// TIA Portal V17 export
// export: Created 2026-11-08T05:50:28.3151889Z, ExportSetting WithDefaults, DisplayName Totally Integrated Automation Portal, DisplayVersion V17, DisplayName TIA Portal Openness, DisplayVersion V17, DisplayName TIA Portal Version Control Interface, DisplayVersion V17, DisplayName STEP 7 Professional, DisplayVersion V17, DisplayName STEP 7 Safety, DisplayVersion V17, DisplayName WinCC Professional, DisplayVersion V17
ORGANIZATION_BLOCK "Main"   // OB1, LAD, ProgramCycle
TITLE = "Main Program Sweep (Cycle)" / Programa principal - Arranque y paro v2
{ S7_Optimized_Access := 'TRUE' }
VERSION : 0.1
// OB1 director: una red por función. Los 3 estilos corren a la vez; el selector de la HMI decide cuál maneja KM1 y los pilotos.
// stored: AutoNumber true, IsIECCheckEnabled false, SetENOAutomatically false
   VAR_INPUT
      Initial_Call : Bool;   // Initial call of this OB
      Remanence : Bool;   // =True, if remanent data are available
   END_VAR
BEGIN

REGION Network 1: MANDO: pulsadores + HMI
   // Une entradas físicas y botones de la HMI.
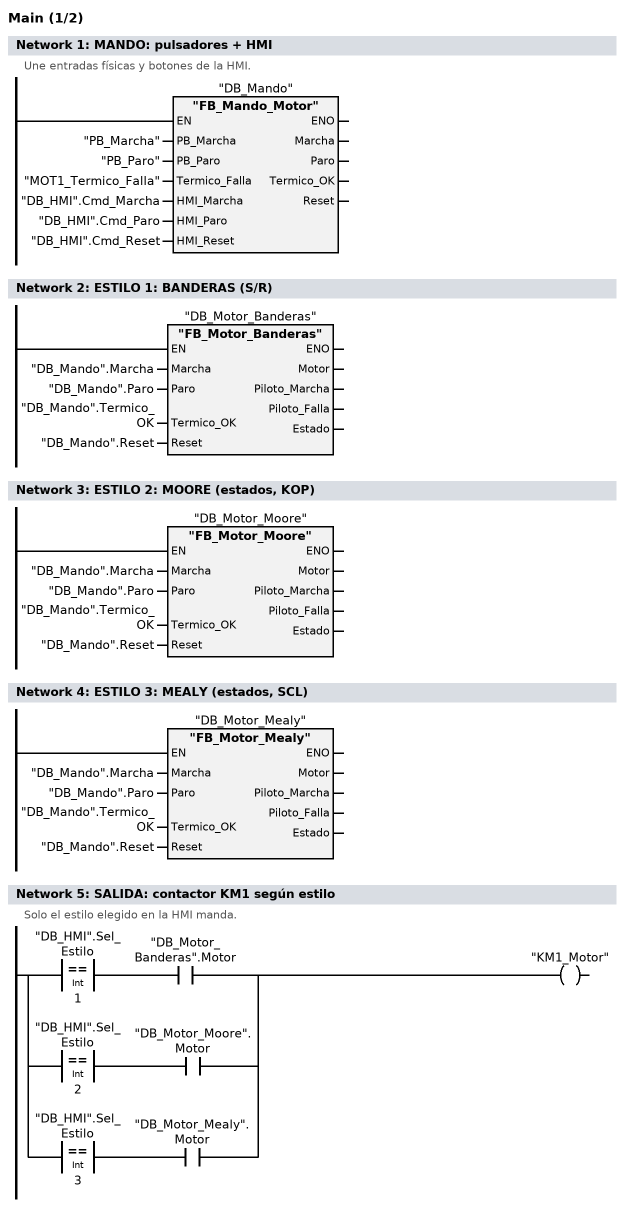
   RUNG wire#powerrail
      "DB_Mando"(PB_Marcha := "PB_Marcha", PB_Paro := "PB_Paro", Termico_Falla := "MOT1_Termico_Falla", HMI_Marcha := "DB_HMI".Cmd_Marcha, HMI_Paro := "DB_HMI".Cmd_Paro, HMI_Reset := "DB_HMI".Cmd_Reset, Marcha =>, Paro =>, Termico_OK =>, Reset =>)
   END_RUNG
   // the same network as SCL:
   "DB_Mando"(PB_Marcha := "PB_Marcha",   // "FB_Mando_Motor"
              PB_Paro := "PB_Paro",
              Termico_Falla := "MOT1_Termico_Falla",
              HMI_Marcha := "DB_HMI".Cmd_Marcha,
              HMI_Paro := "DB_HMI".Cmd_Paro,
              HMI_Reset := "DB_HMI".Cmd_Reset);
END_REGION

REGION Network 2: ESTILO 1: BANDERAS (S/R)
   RUNG wire#powerrail
      "DB_Motor_Banderas"(Marcha := "DB_Mando".Marcha, Paro := "DB_Mando".Paro, Termico_OK := "DB_Mando".Termico_OK, Reset := "DB_Mando".Reset, Motor =>, Piloto_Marcha =>, Piloto_Falla =>, Estado =>)
   END_RUNG
   // the same network as SCL:
   "DB_Motor_Banderas"(Marcha := "DB_Mando".Marcha,   // "FB_Motor_Banderas"
                       Paro := "DB_Mando".Paro,
                       Termico_OK := "DB_Mando".Termico_OK,
                       Reset := "DB_Mando".Reset);
END_REGION

REGION Network 3: ESTILO 2: MOORE (estados, KOP)
   RUNG wire#powerrail
      "DB_Motor_Moore"(Marcha := "DB_Mando".Marcha, Paro := "DB_Mando".Paro, Termico_OK := "DB_Mando".Termico_OK, Reset := "DB_Mando".Reset, Motor =>, Piloto_Marcha =>, Piloto_Falla =>, Estado =>)
   END_RUNG
   // the same network as SCL:
   "DB_Motor_Moore"(Marcha := "DB_Mando".Marcha,   // "FB_Motor_Moore"
                    Paro := "DB_Mando".Paro,
                    Termico_OK := "DB_Mando".Termico_OK,
                    Reset := "DB_Mando".Reset);
END_REGION

REGION Network 4: ESTILO 3: MEALY (estados, SCL)
   RUNG wire#powerrail
      "DB_Motor_Mealy"(Marcha := "DB_Mando".Marcha, Paro := "DB_Mando".Paro, Termico_OK := "DB_Mando".Termico_OK, Reset := "DB_Mando".Reset, Motor =>, Piloto_Marcha =>, Piloto_Falla =>, Estado =>)
   END_RUNG
   // the same network as SCL:
   "DB_Motor_Mealy"(Marcha := "DB_Mando".Marcha,   // "FB_Motor_Mealy"
                    Paro := "DB_Mando".Paro,
                    Termico_OK := "DB_Mando".Termico_OK,
                    Reset := "DB_Mando".Reset);
END_REGION

REGION Network 5: SALIDA: contactor KM1 según estilo
   // Solo el estilo elegido en la HMI manda.
   RUNG wire#powerrail
      { S7_Templates := "SrcType := Int" } EQ_Contact(in1 := "DB_HMI".Sel_Estilo, in2 := 1)
      Contact( "DB_Motor_Banderas".Motor )
      wire#w1
      Coil( "KM1_Motor" )
   END_RUNG
   RUNG wire#powerrail
      { S7_Templates := "SrcType := Int" } EQ_Contact(in1 := "DB_HMI".Sel_Estilo, in2 := 2)
      Contact( "DB_Motor_Moore".Motor )
   END_RUNG wire#w1
   RUNG wire#powerrail
      { S7_Templates := "SrcType := Int" } EQ_Contact(in1 := "DB_HMI".Sel_Estilo, in2 := 3)
      Contact( "DB_Motor_Mealy".Motor )
   END_RUNG wire#w1
   // the same network as SCL:
   "KM1_Motor" := (("DB_HMI".Sel_Estilo = 1) AND "DB_Motor_Banderas".Motor) OR (("DB_HMI".Sel_Estilo = 2) AND "DB_Motor_Moore".Motor) OR (("DB_HMI".Sel_Estilo = 3) AND "DB_Motor_Mealy".Motor);
END_REGION

REGION Network 6: SALIDA: piloto de marcha
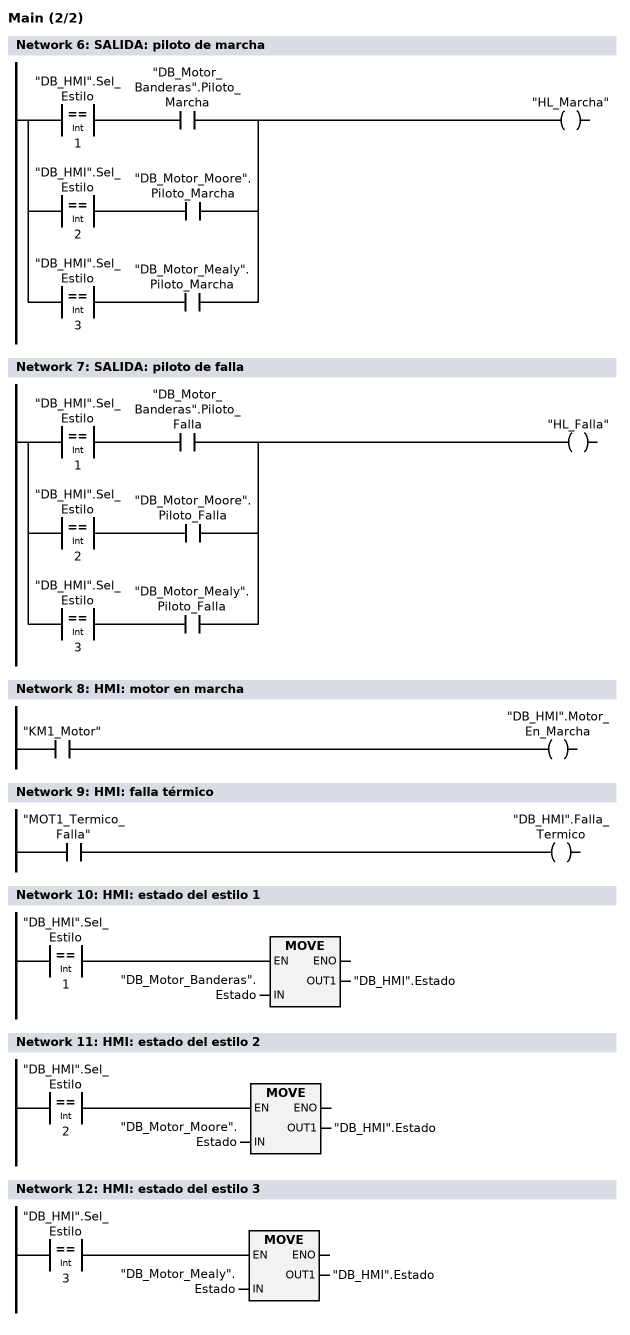
   RUNG wire#powerrail
      { S7_Templates := "SrcType := Int" } EQ_Contact(in1 := "DB_HMI".Sel_Estilo, in2 := 1)
      Contact( "DB_Motor_Banderas".Piloto_Marcha )
      wire#w1
      Coil( "HL_Marcha" )
   END_RUNG
   RUNG wire#powerrail
      { S7_Templates := "SrcType := Int" } EQ_Contact(in1 := "DB_HMI".Sel_Estilo, in2 := 2)
      Contact( "DB_Motor_Moore".Piloto_Marcha )
   END_RUNG wire#w1
   RUNG wire#powerrail
      { S7_Templates := "SrcType := Int" } EQ_Contact(in1 := "DB_HMI".Sel_Estilo, in2 := 3)
      Contact( "DB_Motor_Mealy".Piloto_Marcha )
   END_RUNG wire#w1
   // the same network as SCL:
   "HL_Marcha" := (("DB_HMI".Sel_Estilo = 1) AND "DB_Motor_Banderas".Piloto_Marcha) OR (("DB_HMI".Sel_Estilo = 2) AND "DB_Motor_Moore".Piloto_Marcha) OR (("DB_HMI".Sel_Estilo = 3) AND "DB_Motor_Mealy".Piloto_Marcha);
END_REGION

REGION Network 7: SALIDA: piloto de falla
   RUNG wire#powerrail
      { S7_Templates := "SrcType := Int" } EQ_Contact(in1 := "DB_HMI".Sel_Estilo, in2 := 1)
      Contact( "DB_Motor_Banderas".Piloto_Falla )
      wire#w1
      Coil( "HL_Falla" )
   END_RUNG
   RUNG wire#powerrail
      { S7_Templates := "SrcType := Int" } EQ_Contact(in1 := "DB_HMI".Sel_Estilo, in2 := 2)
      Contact( "DB_Motor_Moore".Piloto_Falla )
   END_RUNG wire#w1
   RUNG wire#powerrail
      { S7_Templates := "SrcType := Int" } EQ_Contact(in1 := "DB_HMI".Sel_Estilo, in2 := 3)
      Contact( "DB_Motor_Mealy".Piloto_Falla )
   END_RUNG wire#w1
   // the same network as SCL:
   "HL_Falla" := (("DB_HMI".Sel_Estilo = 1) AND "DB_Motor_Banderas".Piloto_Falla) OR (("DB_HMI".Sel_Estilo = 2) AND "DB_Motor_Moore".Piloto_Falla) OR (("DB_HMI".Sel_Estilo = 3) AND "DB_Motor_Mealy".Piloto_Falla);
END_REGION

REGION Network 8: HMI: motor en marcha
   RUNG wire#powerrail
      Contact( "KM1_Motor" )
      Coil( "DB_HMI".Motor_En_Marcha )
   END_RUNG
   // the same network as SCL:
   "DB_HMI".Motor_En_Marcha := "KM1_Motor";
END_REGION

REGION Network 9: HMI: falla térmico
   RUNG wire#powerrail
      Contact( "MOT1_Termico_Falla" )
      Coil( "DB_HMI".Falla_Termico )
   END_RUNG
   // the same network as SCL:
   "DB_HMI".Falla_Termico := "MOT1_Termico_Falla";
END_REGION

REGION Network 10: HMI: estado del estilo 1
   RUNG wire#powerrail
      { S7_Templates := "SrcType := Int" } EQ_Contact(in1 := "DB_HMI".Sel_Estilo, in2 := 1)
      { S7_GenerateENO := "TRUE" } Move(in := "DB_Motor_Banderas".Estado, out1 => "DB_HMI".Estado)
   END_RUNG
   // the same network as SCL:
   IF "DB_HMI".Sel_Estilo = 1 THEN "DB_HMI".Estado := "DB_Motor_Banderas".Estado; END_IF;
END_REGION

REGION Network 11: HMI: estado del estilo 2
   RUNG wire#powerrail
      { S7_Templates := "SrcType := Int" } EQ_Contact(in1 := "DB_HMI".Sel_Estilo, in2 := 2)
      { S7_GenerateENO := "TRUE" } Move(in := "DB_Motor_Moore".Estado, out1 => "DB_HMI".Estado)
   END_RUNG
   // the same network as SCL:
   IF "DB_HMI".Sel_Estilo = 2 THEN "DB_HMI".Estado := "DB_Motor_Moore".Estado; END_IF;
END_REGION

REGION Network 12: HMI: estado del estilo 3
   RUNG wire#powerrail
      { S7_Templates := "SrcType := Int" } EQ_Contact(in1 := "DB_HMI".Sel_Estilo, in2 := 3)
      { S7_GenerateENO := "TRUE" } Move(in := "DB_Motor_Mealy".Estado, out1 => "DB_HMI".Estado)
   END_RUNG
   // the same network as SCL:
   IF "DB_HMI".Sel_Estilo = 3 THEN "DB_HMI".Estado := "DB_Motor_Mealy".Estado; END_IF;
END_REGION
END_ORGANIZATION_BLOCK
